// TIA Portal V20 export
// export: Created 2026-10-12T16:46:20.8888353Z, ExportSetting WithDefaults, DisplayName Totally Integrated Automation Portal, DisplayVersion V20 Update 6, DisplayName TIA Portal Openness, DisplayVersion V20 Update 6, DisplayName TIA Portal Version Control Interface, DisplayVersion V20 Update 6, DisplayName SINAMICS Startdrive Advanced, DisplayVersion V20 SP1 Update 2, DisplayName SINAMICS Startdrive G110M, G120, G120C, G120D, G120P, G115D, DisplayVersion V20 SP1 Update 2, DisplayName SINAMICS Startdrive G130, G150, S120, S150, SINAMICS MV, G220, S200, S210, DisplayVersion V20 SP1 Update 2, DisplayName STEP 7 Professional, DisplayVersion V20 Update 6, DisplayName STEP 7 Safety, DisplayVersion V20 Update 2, DisplayName WinCC Basic/Comfort/Advanced, DisplayVersion V20 Update 6, DisplayName WinCC Professional, DisplayVersion V20 Update 6, DisplayName WinCC Unified, DisplayVersion V20 Update 6
FUNCTION_BLOCK "FB_Heizungsregelung"   // FB10, SCL
{ S7_Optimized_Access := 'TRUE' }
VERSION : 0.1
// stored: AutoNumber true, IsIECCheckEnabled false, IsRetainMemResEnabled false, MemoryReserve 100, SetENOAutomatically false, UDAEnableTagReadback false
   VAR_INPUT
      Soll : Real;
      Ist : Real;
      Freigabe : Bool;
   END_VAR
   VAR_OUTPUT
      Schuetz : Bool;
      PT100_Stoerung : Bool;
   END_VAR
   VAR
      Schuetz_Intern : Bool;
   END_VAR
   VAR_TEMP
      einschaltSchwelle : Real;
      ausschaltSchwelle : Real;
   END_VAR
   VAR CONSTANT
      HYSTERESE : Real := 0.2;
      PT100_MIN : Real := -10.0;
      PT100_MAX : Real := 200.0;
   END_VAR
BEGIN

       #PT100_Stoerung:=(#Ist<#PT100_MIN)OR(#Ist>#PT100_MAX);
       IF NOT #Freigabe OR(#Soll<=0.0)OR #PT100_Stoerung THEN #Schuetz_Intern:=FALSE; #Schuetz:=FALSE; RETURN; END_IF;
       #einschaltSchwelle:=#Soll-(#HYSTERESE/2.0); #ausschaltSchwelle:=#Soll+(#HYSTERESE/2.0);
       IF #Ist<#einschaltSchwelle THEN #Schuetz_Intern:=TRUE; ELSIF #Ist>#ausschaltSchwelle THEN #Schuetz_Intern:=FALSE; END_IF;
       #Schuetz:=#Schuetz_Intern;
END_FUNCTION_BLOCK
